SUBAPPLICATION GreenRedBackground4SC (* Hintergrundfarbe (TRUE -> Grün, FALSE -> Rot) für 4 Objekte (Kompakt) *)
  (* Standard: 61499-2 *)
  (* Version 1.0, 2026-07-21, franz, Meisterschulen am Ostbahnhof *)
  PACKAGE MyLib::sys;
  IMPORT isobus::UT::Q::types::s3ObjectIDs;
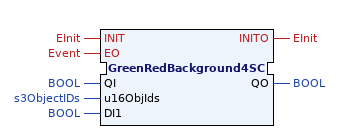
  EVENT_INPUT
    INIT : EInit; (* Initialization Request *)
    EO;
  END_EVENT
  EVENT_OUTPUT
    INITO : EInit; (* Initialization Confirm *)
  END_EVENT
  VAR_INPUT
    QI : BOOL := TRUE; (* Quality Input - TRUE to enable service *)
    u16ObjIds : isobus::UT::Q::types::s3ObjectIDs;
    DI1 : BOOL; (* Selector *)
  END_VAR
  VAR_OUTPUT
    QO : BOOL; (* Quality Output - TRUE if service executed successfully *)
  END_VAR
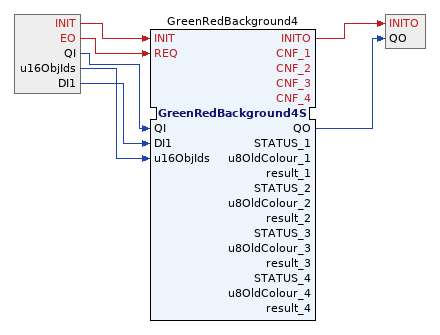
  SUBAPPS
    GreenRedBackground4 : MyLib::sys::GreenRedBackground4S;
  END_SUBAPPS
  EVENT_CONNECTIONS
    EO TO GreenRedBackground4.REQ;
    INIT TO GreenRedBackground4.INIT;
    GreenRedBackground4.INITO TO INITO;
  END_CONNECTIONS
  DATA_CONNECTIONS
    u16ObjIds TO GreenRedBackground4.u16ObjIds;
    DI1 TO GreenRedBackground4.DI1;
    QI TO GreenRedBackground4.QI;
    GreenRedBackground4.QO TO QO;
  END_CONNECTIONS
END_SUBAPPLICATION
